(*
SPDX-FileCopyrightText: © 2026 Oleksandr Tiutyk <trofimich@gmail.com>
SPDX-License-Identifier: MIT
License: https://opensource.org/license/mit
*)

(*!
<summary>
Named variable lookup reports failure without propagating exceptions; its output is usable only on success.
</summary>
*)
INTERFACE IVariableLookup EXTENDS TOF_Core.IObject

(*!
<summary>Attempts to resolve a named variable from the available variable containers.</summary>
<description>
Returns FALSE when resolution fails or a nested call raises an exception. Use the output only when TRUE is
returned. Does not propagate exceptions or clear terminal allocation state. Terminal allocation failure forces FALSE,
including when a nested lookup contained its original exception. The owner still raises at the task boundary.
</description>
<param name="name">Case-sensitive variable name to resolve.</param>
<param name="variable">Borrowed generic value descriptor on TRUE; unassigned on FALSE.</param>
*)
METHOD TryGetVariable : BOOL
VAR_INPUT
	name : STRING;
END_VAR
VAR_OUTPUT
	variable : TOF_Core.GENERIC_VALUE;
END_VAR
END_METHOD

END_INTERFACE

(* stored: Version 1.1.0.1
   Itf IVariableLookup: Id {9265c155-6fb7-43aa-a2f1-419ffde75d0d}
   Method TryGetVariable: Id {473aa1d0-5468-4e6f-b2a4-5c756ab0236e} *)
